NAMESPACE TiaMcp_UnitA.Alternate
FUNCTION_BLOCK "TgpNamespace_NestEffect"
{ S7_Optimized_Access := 'TRUE' }
VERSION : 0.1
VAR_INPUT
 Enable : Bool;
END_VAR
VAR_OUTPUT
 Active : Bool;
END_VAR
VAR
 RetainedMarker : Int := 17;
END_VAR
BEGIN
 #Active := #Enable;
END_FUNCTION_BLOCK

FUNCTION_BLOCK "TgpNamespace_NestParent"
{ S7_Optimized_Access := 'TRUE' }
VERSION : 0.1
VAR_INPUT
 Enable : Bool;
END_VAR
VAR_OUTPUT
 Active : Bool;
END_VAR
VAR
 RetainedMarker : Int := 17;
 Inner : "TiaMcp_UnitA.Alternate.TgpNamespace_NestEffect";
END_VAR
BEGIN
 #Active := #Enable;
END_FUNCTION_BLOCK

FUNCTION_BLOCK "TgpNamespace_NestGrand"
{ S7_Optimized_Access := 'TRUE' }
VERSION : 0.1
VAR_INPUT
 Enable : Bool;
END_VAR
VAR_OUTPUT
 Active : Bool;
END_VAR
VAR
 RetainedMarker : Int := 17;
 Middle : "TiaMcp_UnitA.Alternate.TgpNamespace_NestParent";
END_VAR
BEGIN
 #Active := #Enable;
END_FUNCTION_BLOCK

DATA_BLOCK "TgpNamespace_NestEffect_DB"
{ S7_Optimized_Access := 'TRUE' }
VERSION : 0.1
"TiaMcp_UnitA.Alternate.TgpNamespace_NestEffect"
BEGIN
 RetainedMarker := 42;
END_DATA_BLOCK

DATA_BLOCK "TgpNamespace_NestParent_DB"
{ S7_Optimized_Access := 'TRUE' }
VERSION : 0.1
"TiaMcp_UnitA.Alternate.TgpNamespace_NestParent"
BEGIN
 RetainedMarker := 42;
 Inner.RetainedMarker := 42;
END_DATA_BLOCK

DATA_BLOCK "TgpNamespace_NestGrand_DB"
{ S7_Optimized_Access := 'TRUE' }
VERSION : 0.1
"TiaMcp_UnitA.Alternate.TgpNamespace_NestGrand"
BEGIN
 RetainedMarker := 42;
 Middle.RetainedMarker := 42;
 Middle.Inner.RetainedMarker := 42;
END_DATA_BLOCK

END_NAMESPACE
